RoboDK station: first project.rdk

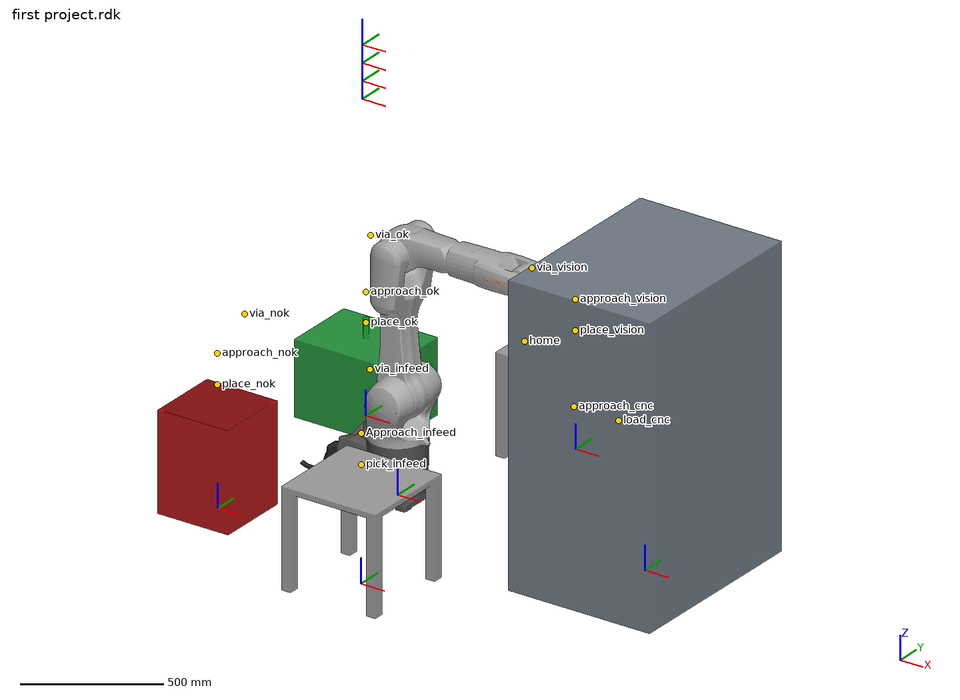
[picture v0: the station drawn from its stored meshes, robots at their saved joint values, targets as dots, program paths as lines]
Station KUKA_Cell (saved by RoboDK 6.1.1). Poses are relative to the parent item; angles as X-Y-Z fixed-axis rotations.
  - frame KUKA KR 10 R1100-2 Base at (0, 0, 0) mm
    - robot KUKA KR 10 R1100-2: 6 axes, payload 10.9 kg, reach 1101 mm, repeatability 0.02 mm, weight 56.5 kg
        modified DH rows (alpha deg, a mm, theta deg, d mm): 0, 0, 0, 400; -90, 25, 0, 0; 0, 560, -90, 0; -90, 25, 0, 515; 90, 0, 0, 0; -90, 0, 180, 90
        joint limits [-170, -190, -120, -185, -120, -350] to [170, 45, 156, 185, 120, 350]; home [0, -90, 90, 0, 0, 0]; saved at [0, -90, 90, 0, 90, 0]
      - tool Tool_Gripper, TCP at (0, 0, 150) mm, size 90 x 80 x 150 mm
    - target home (joint target) at (540, 0, 745) mm, rotated rx 180 ry 0 rz -180 deg; joints [0, -90, 90, 0, 90, 0] of KUKA KR 10 R1100-2
    - target via_infeed (joint target) at (226.29, -490.3, 745) mm, rotated rx 180 ry 0 rz 114.78 deg; joints [65.225, -90, 90, 0, 90, 0] of KUKA KR 10 R1100-2
    - target via_cnc (joint target) at (540, 0, 745) mm, rotated rx 180 ry 0 rz -180 deg; joints [0, -90, 90, 0, 90, 0] of KUKA KR 10 R1100-2
    - target via_vision (joint target) at (226.29, 490.3, 745) mm, rotated rx 180 ry 0 rz -114.78 deg; joints [-65.225, -90, 90, 0, 90, 0] of KUKA KR 10 R1100-2
    - target via_ok (joint target) at (-381.84, 381.84, 745) mm, rotated rx 180 ry 0 rz -45 deg; joints [-135, -90, 90, 0, 90, 0] of KUKA KR 10 R1100-2
    - target via_nok (joint target) at (-381.84, -381.84, 745) mm, rotated rx 180 ry 0 rz 45 deg; joints [135, -90, 90, 0, 90, 0] of KUKA KR 10 R1100-2
  - Python program check_paths (listed below)
  - Python program main_cycle (1) (listed below)
  - Python program build_cell (1) (listed below)
  - frame Frame_Infeed at (300, -650, 0) mm
    - object Table_Infeed at (0, 0, 0) mm, size 400 x 400 x 400 mm, geometry from Table.stl
    - target Approach_infeed (Cartesian target) at (0, 0, 580) mm, rotated rx 180 ry 0 rz 0 deg; joints [65.225, -70.524, 85.389, 0, 75.135, -114.775] of KUKA KR 10 R1100-2
    - target pick_infeed (Cartesian target) at (0, 0, 460) mm, rotated rx 180 ry 0 rz 0 deg; joints [65.225, -66.659, 93.982, 0, 62.678, -114.775] of KUKA KR 10 R1100-2
  - frame Frame_CNC at (1050, 0, 0) mm
    - object CNC_Machine at (0, 0, 0) mm, size 600 x 800 x 1200 mm, geometry from CNC_Machine.stl
    - target approach_cnc (Cartesian target) at (-300, 0, 550) mm, rotated rx 0 ry 90 rz 0 deg; joints [0, -74.689, 126.636, 0, -51.947, 0] of KUKA KR 10 R1100-2
    - target load_cnc (Cartesian target) at (-110, 0, 550) mm, rotated rx 0 ry 90 rz 0 deg; joints [0, -59.76, 102.885, 0, -43.124, 0] of KUKA KR 10 R1100-2
  - frame Frame_Vision at (300, 650, 0) mm
    - object Table_Vision at (0, 0, 0) mm, size 400 x 400 x 400 mm, geometry from Table.stl
    - target approach_vision (Cartesian target) at (0, 0, 580) mm, rotated rx 180 ry 0 rz 0 deg; joints [-65.225, -70.524, 85.389, 0, 75.135, 114.775] of KUKA KR 10 R1100-2
    - target place_vision (Cartesian target) at (0, 0, 460) mm, rotated rx 180 ry 0 rz 0 deg; joints [-65.225, -66.659, 93.982, 0, 62.678, 114.775] of KUKA KR 10 R1100-2
  - frame Frame_OK at (-450, 450, 0) mm
    - object Pallet_OK at (0, 0, 0) mm, size 400 x 300 x 300 mm, geometry from Pallet_OK.stl
    - target approach_ok (Cartesian target) at (0, 0, 480) mm, rotated rx 180 ry 0 rz 0 deg; joints [-135, -74.946, 103.078, 0, 61.868, 45] of KUKA KR 10 R1100-2
    - target place_ok (Cartesian target) at (0, 0, 360) mm, rotated rx 180 ry 0 rz 0 deg; joints [-135, -68.275, 109.448, 0, 48.827, 45] of KUKA KR 10 R1100-2
    - object Part_Shaft at (0, 0, 300) mm, size 20 x 20 x 80 mm, geometry from Part_Shaft.stl
  - frame Frame_NOK at (-450, -450, 0) mm
    - object Bin_NOK at (0, 0, 0) mm, size 300 x 300 x 400 mm, geometry from Bin_NOK.stl
    - target approach_nok (Cartesian target) at (0, 0, 600) mm, rotated rx 180 ry 0 rz 0 deg; joints [135, -78.926, 93.974, 0, 74.951, -45] of KUKA KR 10 R1100-2
    - target place_nok (Cartesian target) at (0, 0, 480) mm, rotated rx 180 ry 0 rz 0 deg; joints [135, -74.946, 103.078, 0, 61.868, -45] of KUKA KR 10 R1100-2
  - Python program kpi_report (listed below)
  - Python program dashboard (listed below)
  - frame HMI | ORDER OF-20261010-1825: 5 parts  |  now: SN-0005 at (-150, 0, 1700) mm
  - frame HMI | Status: ORDER FINISHED at (-150, 0, 1630) mm
  - frame HMI | Last: SN-0005  D=20.005 mm  OK  11.5 s  stop 152 s at (-150, 0, 1560) mm
  - frame HMI | Done 5/5   OK: 5   NOK: 0   Yield: 100 %   Downtime: 240 s at (-150, 0, 1490) mm

--- Python program check_paths ---
# =====================================================================
#  check_paths.py  -  checks every robot move of the cycle
#
#  For each move it checks:
#    1. REACH      : the robot can reach the target
#    2. COLLISION  : no collision along the path (robot / gripper vs cell)
#    3. LINEAR     : the straight-line (LIN) move is possible
#    4. SINGULARITY: wrist A5 not close to 0 deg (KUKA wrist singularity)
#    5. JOINT LIMIT: no joint closer than 5 deg to its limit
#
#  Run main_cycle.py at least once before (it writes the target values).
#  Result: a report in RoboDK + path_check_report.csv next to the station.
# =====================================================================
import csv
import os

from robodk.robolink import (Robolink, ITEM_TYPE_ROBOT, ITEM_TYPE_TOOL, ITEM_TYPE_TARGET,
                             ITEM_TYPE_FRAME, ITEM_TYPE_OBJECT, COLLISION_ON, COLLISION_OFF)
from robodk.robomath import transl

RDK = Robolink()

SIM_SPEED = 1          # 1 = real speed (slow, easy to watch). 5 = faster
SINGULARITY_DEG = 10   # warn if |A5| below this
LIMIT_MARGIN_DEG = 5   # warn if a joint is this close to its limit
HOME_JOINTS = [0, -90, 90, 0, 90, 0]

def find_robot_and_tool():
    """KUKA robot (ignores a gripper mechanism) + its gripper tool."""
    robots = RDK.ItemList(ITEM_TYPE_ROBOT)
    if not robots:
        raise Exception("No robot in the station. Load the KUKA KR 10 first.")
    rob = next((r for r in robots if "KUKA" in r.Name().upper()), robots[0])
    tl = RDK.Item('Tool_Gripper', ITEM_TYPE_TOOL)
    if not tl.Valid() or tl.Name() != 'Tool_Gripper':
        tools = [t for t in RDK.ItemList(ITEM_TYPE_TOOL)]
        if not tools:
            tl = rob.AddTool(transl(0, 0, 150), 'Tool_Gripper')
        else:
            tl = tools[0]
            tl.setName('Tool_Gripper')
    return rob, tl


robot, tool = find_robot_and_tool()
part = RDK.Item('Part_Shaft', ITEM_TYPE_OBJECT)
robot.setPoseTool(tool)


def collision_report():
    """Names of the items that are touching right now (empty string if none)."""
    try:
        pairs = RDK.CollisionPairs()            # [[item1, item2, link1, link2], ...]
        out = []
        for p in pairs:
            a = p[0].Name() + (f" (J{p[2]})" if len(p) > 2 and p[0].Type() == ITEM_TYPE_ROBOT else "")
            b = p[1].Name() + (f" (J{p[3]})" if len(p) > 3 and p[1].Type() == ITEM_TYPE_ROBOT else "")
            out.append(f"{a}  <->  {b}")
        return "; ".join(out)
    except Exception:
        try:
            return ", ".join(i.Name() for i in RDK.CollisionItems())
        except Exception:
            return ""


def choose_home():
    """Pick the home where the gripper points DOWN (A5 = +90 or -90).
    A home with the gripper pointing up makes the wrist flip during the moves
    and the gripper fingers hit the robot arm (self-collision)."""
    global HOME_JOINTS
    for a5 in (90, -90):
        j = [0, -90, 90, 0, a5, 0]
        robot.setJoints(j)
        tcp = robot.Pose()                  # TCP pose (active tool) in robot base
        if tcp[2, 2] < -0.5:                # tool Z axis points down
            HOME_JOINTS = j
            print(f"Home: A5 = {a5} (gripper pointing down)")
            return j
    return HOME_JOINTS

# Same sequence as main_cycle (OK branch + NOK branch)
SEQUENCE = [
    ("J", "home"),
    ("J", "via_infeed"), ("J", "Approach_infeed"), ("L", "pick_infeed"), ("GRIP", None),
    ("L", "Approach_infeed"), ("J", "via_infeed"),
    ("J", "via_cnc"), ("J", "approach_cnc"), ("L", "load_cnc"), ("RELEASE", "Frame_CNC"),
    ("L", "approach_cnc"), ("L", "load_cnc"), ("GRIP", None), ("L", "approach_cnc"), ("J", "via_cnc"),
    ("J", "via_vision"), ("J", "approach_vision"), ("L", "place_vision"), ("RELEASE", "Frame_Vision"),
    ("L", "approach_vision"), ("L", "place_vision"), ("GRIP", None), ("L", "approach_vision"),
    ("J", "via_vision"),
    ("J", "via_ok"), ("J", "approach_ok"), ("L", "place_ok"), ("RELEASE", "Frame_OK"),
    ("L", "approach_ok"), ("J", "via_ok"),
    ("J", "via_nok"), ("J", "approach_nok"), ("L", "place_nok"), ("L", "approach_nok"),  # NOK (empty gripper)
    ("J", "via_nok"),
    ("J", "home"),
]


def item(name, itype):
    it = RDK.Item(name, itype)
    if not it.Valid():
        raise Exception(f"Not found in the tree: {name}")
    return it


def disable_part_collisions():
    """The part touches the gripper and tables on purpose -> ignore it."""
    for other in RDK.ItemList():
        for link in range(8):
            try:
                RDK.setCollisionActivePair(COLLISION_OFF, part, other, 0, link)
            except Exception:
                pass


def as_list(values):
    """RoboDK returns joints as a Mat object -> convert to a flat Python list."""
    if hasattr(values, "rows"):          # robodk Mat (column or row vector)
        values = values.rows
    elif hasattr(values, "list"):
        values = values.list()
    out = []
    for v in values:
        if isinstance(v, (list, tuple)):
            out.extend(v)
        else:
            out.append(v)
    return [float(x) for x in out]


def check_joints(joints):
    """Return a list of warnings for singularity and joint limits."""
    warnings = []
    j = as_list(joints)
    if len(j) < 6:
        return warnings
    if abs(j[4]) < SINGULARITY_DEG:
        warnings.append(f"A5={j[4]:.1f} deg (near singularity)")
    limits = robot.JointLimits()
    lower, upper = as_list(limits[0]), as_list(limits[1])
    for i in range(6):
        if j[i] - lower[i] < LIMIT_MARGIN_DEG or upper[i] - j[i] < LIMIT_MARGIN_DEG:
            warnings.append(f"A{i+1}={j[i]:.1f} deg (near limit)")
    return warnings


# ---------------------------------------------------------------- run
RDK.setSimulationSpeed(SIM_SPEED)
RDK.setCollisionActive(COLLISION_ON)
disable_part_collisions()

part.setParent(item('Frame_Infeed', ITEM_TYPE_FRAME))
part.setPose(transl(0, 0, 400))
via = RDK.Item('via_infeed', ITEM_TYPE_TARGET)
if not via.Valid() or via.Name() != 'via_infeed':
    raise Exception('Run main_cycle once first (it creates the via_ points).')
robot.setJoints(item('home', ITEM_TYPE_TARGET).Joints())

report = []
n_problems = 0

for step, (kind, name) in enumerate(SEQUENCE, start=1):
    if kind == "GRIP":
        part.setParentStatic(tool)
        continue
    if kind == "RELEASE":
        part.setParentStatic(item(name, ITEM_TYPE_FRAME))
        continue

    target = item(name, ITEM_TYPE_TARGET)
    j_start = robot.Joints()
    row = {"step": step, "move": "PTP" if kind == "J" else "LIN", "target": name,
           "reach": "OK", "linear": "-", "collisions": 0, "hit": "", "warnings": "", "status": "OK"}

    # Test LIN feasibility before moving
    if kind == "L":
        robot.setPoseFrame(target.Parent())
        res = robot.MoveL_Test(j_start, target.Pose())
        row["linear"] = "OK" if res == 0 else ("collision" if res > 0 else "NOT POSSIBLE")

    # Execute the move (PTP if LIN impossible, like main_cycle does)
    try:
        if kind == "L" and row["linear"] != "NOT POSSIBLE":
            robot.MoveL(target)
        else:
            robot.MoveJ(target.Joints())     # joints computed by main_cycle setup
    except Exception:
        row["reach"] = "STOPPED (collision or unreachable)"
        row["hit"] = collision_report()
        row["status"] = "FAIL"
        report.append(row)
        n_problems += 1
        print(f"{step:02d} {name:16s} STOPPED (collision or unreachable)")
        break

    j_end = robot.Joints()
    # Collision along the joint path (PTP) or at the end pose
    if kind == "J":
        row["collisions"] = max(0, robot.MoveJ_Test(j_start, j_end))
    else:
        row["collisions"] = max(0, RDK.Collisions())
    if row["collisions"] > 0:
        row["hit"] = collision_report()
    warnings = check_joints(j_end)
    row["warnings"] = "; ".join(warnings)

    if row["collisions"] > 0 or row["linear"] in ("collision", "NOT POSSIBLE"):
        row["status"] = "FAIL"
    elif warnings:
        row["status"] = "WARNING"
    if row["status"] != "OK":
        n_problems += 1

    report.append(row)
    print(f"{step:02d} {row['move']} {name:16s} reach={row['reach']:4s} "
          f"lin={row['linear']:12s} coll={row['collisions']} {row['status']} {row['warnings']}")

RDK.setCollisionActive(COLLISION_OFF)

# ---------------------------------------------------------------- report
station_path = RDK.getParam('PATH_OPENSTATION')
out_dir = station_path if station_path and os.path.isdir(station_path) else os.path.expanduser("~")
out_file = os.path.join(out_dir, "path_check_report.csv")
with open(out_file, "w", newline="") as f:
    w = csv.DictWriter(f, fieldnames=list(report[0].keys()))
    w.writeheader()
    w.writerows(report)

lines = [f"{r['step']:02d} {r['move']} {r['target']}: {r['status']}"
         + (f" {r['reach']}" if r['reach'] != 'OK' else "")
         + (f" ({r['warnings']})" if r['warnings'] else "")
         + (f" collisions={r['collisions']}" if r['collisions'] else "")
         + (f"\n      HIT: {r['hit']}" if r['hit'] else "")
         + (f" LIN={r['linear']}" if r['linear'] not in ('-', 'OK') else "")
         for r in report]
summary = ("ALL PATHS OK" if n_problems == 0 else f"{n_problems} PROBLEM(S) FOUND")
RDK.ShowMessage(summary + "\n\n" + "\n".join(lines) + f"\n\nReport: {out_file}", True)
print(summary, "->", out_file)

--- Python program main_cycle (1) ---
# =====================================================================
#  KUKA KR 10 machine-tending cell - main cycle (RoboDK Python API)
#
#  1. SETUP : writes every target, picks ONE consistent arm configuration
#             per station (no wrist flips) and creates a safe "via" point
#             above each station.
#  2. CYCLE : pick -> CNC -> vision -> OK / NOK, always moving between
#             stations at safe height (via points).
#  3. LOG   : one CSV line per part (for the MES dashboard).
#
#  Tip: run it once with collision checking OFF (setup), then check_paths.
# =====================================================================
import csv
import math
import os
import random
import time
from datetime import datetime

from robodk.robolink import (Robolink, ITEM_TYPE_ROBOT, ITEM_TYPE_TOOL,
                             ITEM_TYPE_TARGET, ITEM_TYPE_FRAME, ITEM_TYPE_OBJECT,
                             COLLISION_ON, COLLISION_OFF)
from robodk.robomath import transl, invH, KUKA_2_Pose

RDK = Robolink()

# ---------------------------------------------------------------- settings
N_PARTS = 5                      # number of parts to produce
MACHINING_TIME_S = 3             # simulated CNC cycle
NOMINAL_DIAM = 20.00             # mm
TOLERANCE = 0.05                 # mm  -> OK if 19.95 .. 20.05
_station_dir = RDK.getParam('PATH_OPENSTATION')          # folder of the saved station
LOG_DIR = _station_dir if _station_dir and os.path.isdir(str(_station_dir)) else \
    os.path.join(os.path.expanduser("~"), "Documents", "KUKA_Cell_MES")
LOG_FILE = os.path.join(LOG_DIR, "kuka_cell_log.csv")   # CSV saved next to KUKA_Cell.rdk
CNC_FRAME_X = 1050               # CNC farther: more space between robot and CNC door

# ---------------------------------------------------------------- STEP 1: faults & downtime
# Each fault: (station, stop reason, probability per part, min-max stop duration in seconds)
FAULTS = [
    ("infeed", "Part missing on infeed",   0.10, (20, 60)),
    ("infeed", "Gripper fault",            0.05, (30, 90)),
    ("cnc",    "CNC door not open",        0.08, (15, 45)),
    ("cnc",    "Tool change on CNC",       0.05, (60, 180)),
    ("vision", "Camera timeout",           0.07, (10, 30)),
]
TIME_SCALE = 0.05                # a 60 s stop is shown as 3 s in the simulation
EVENT_FILE = os.path.join(LOG_DIR, "kuka_cell_events.csv")   # one line per stop
ORDER_ID = datetime.now().strftime("OF-%Y%m%d-%H%M")         # production order number

# Stations: name -> (frame, approach target, work target, approach values, work values)
# values = (X, Y, Z, A=rz, B=ry, C=rx) in the station frame (KUKA convention)
STATIONS = {
    "infeed": ("Frame_Infeed", "Approach_infeed", "pick_infeed",
               (0, 0, 580, 0, 0, 180), (0, 0, 460, 0, 0, 180)),
    "cnc":    ("Frame_CNC", "approach_cnc", "load_cnc",
               (-300, 0, 550, 0, 90, 0), (-110, 0, 550, 0, 90, 0)),
    "vision": ("Frame_Vision", "approach_vision", "place_vision",
               (0, 0, 580, 0, 0, 180), (0, 0, 460, 0, 0, 180)),
    "ok":     ("Frame_OK", "approach_ok", "place_ok",
               (0, 0, 480, 0, 0, 180), (0, 0, 360, 0, 0, 180)),
    "nok":    ("Frame_NOK", "approach_nok", "place_nok",
               (0, 0, 600, 0, 0, 180), (0, 0, 480, 0, 0, 180)),
}
HOME_JOINTS = [0, -90, 90, 0, 90, 0]
SOLVED = {}        # target name -> joints computed in setup (used by MoveJ)

# ---------------------------------------------------------------- items
def find_robot_and_tool():
    """KUKA robot (ignores a gripper mechanism) + its gripper tool."""
    robots = RDK.ItemList(ITEM_TYPE_ROBOT)
    if not robots:
        raise Exception("No robot in the station. Load the KUKA KR 10 first.")
    rob = next((r for r in robots if "KUKA" in r.Name().upper()), robots[0])
    tl = RDK.Item('Tool_Gripper', ITEM_TYPE_TOOL)
    if not tl.Valid() or tl.Name() != 'Tool_Gripper':
        tools = [t for t in RDK.ItemList(ITEM_TYPE_TOOL)]
        if not tools:
            tl = rob.AddTool(transl(0, 0, 150), 'Tool_Gripper')
        else:
            tl = tools[0]
            tl.setName('Tool_Gripper')
    return rob, tl


robot, tool = find_robot_and_tool()
part = RDK.Item('Part_Shaft', ITEM_TYPE_OBJECT)
robot.setPoseTool(tool)


def collision_report():
    """Names of the items that are touching right now (empty string if none)."""
    try:
        pairs = RDK.CollisionPairs()            # [[item1, item2, link1, link2], ...]
        out = []
        for p in pairs:
            a = p[0].Name() + (f" (J{p[2]})" if len(p) > 2 and p[0].Type() == ITEM_TYPE_ROBOT else "")
            b = p[1].Name() + (f" (J{p[3]})" if len(p) > 3 and p[1].Type() == ITEM_TYPE_ROBOT else "")
            out.append(f"{a}  <->  {b}")
        return "; ".join(out)
    except Exception:
        try:
            return ", ".join(i.Name() for i in RDK.CollisionItems())
        except Exception:
            return ""
robot.setPoseFrame(robot.Parent())      # poses measured in the robot base


def T(name):
    item = RDK.Item(name, ITEM_TYPE_TARGET)
    if not item.Valid() or item.Name() != name:
        raise Exception(f"Target not found in the tree: {name}")
    return item


def F(name):
    item = RDK.Item(name, ITEM_TYPE_FRAME)
    if not item.Valid():
        raise Exception(f"Frame not found in the tree: {name}")
    return item


def as_list(values):
    """RoboDK returns joints as a Mat -> flat Python list."""
    if hasattr(values, "rows"):
        values = values.rows
    elif hasattr(values, "list"):
        values = values.list()
    out = []
    for v in values:
        out.extend(v) if isinstance(v, (list, tuple)) else out.append(v)
    return [float(x) for x in out]


# ---------------------------------------------------------------- moves
def MJ(name):
    try:
        if name in SOLVED:
            robot.MoveJ(SOLVED[name])        # exact joints from setup: no config surprise
        else:
            robot.MoveJ(T(name))
    except Exception as e:
        hit = collision_report()
        msg = f"Move stopped going to: {name}" + (f"\nCOLLISION: {hit}" if hit else f" ({e})")
        RDK.ShowMessage(msg, True)
        raise Exception(msg)


def ML(name):
    try:
        robot.MoveL(T(name))
    except Exception:
        print(f"  MoveL to {name} not possible -> MoveJ used")
        MJ(name)


def grip():
    part.setParentStatic(tool)


def release(frame_name):
    part.setParentStatic(F(frame_name))


# ---------------------------------------------------------------- on-screen display (HMI)
# RoboDK shows the NAME of a frame as a text label in the 3D view.
# We create 4 small frames above the cell and change their names = live text panel.
HMI_POS = (-150, 0, 1700)          # where the text panel floats (mm, station frame)
HMI = []
PART_COLOR = [0.85, 0.65, 0.20, 1]   # gold = raw part


def hmi_init():
    for fr in RDK.ItemList(ITEM_TYPE_FRAME):          # remove the panel of a previous run
        if fr.Name().startswith("HMI"):
            fr.Delete()
    HMI.clear()
    for i in range(4):
        fr = RDK.AddFrame(f"HMI {i}")
        fr.setPose(transl(HMI_POS[0], HMI_POS[1], HMI_POS[2] - 70 * i))
        try:
            fr.setVisible(True, False)                  # show the text, hide the axes
        except Exception:
            pass
        HMI.append(fr)


def hmi(line, text):
    """Write one line of the 3D text panel (0 = title, 1 = status, 2 = last part, 3 = totals)."""
    if line < len(HMI):
        HMI[line].setName(f"HMI | {text}")


def color_part(rgba):
    try:
        part.setColor(rgba)
    except Exception:
        pass


def reset_part():
    part.setParent(F('Frame_Infeed'))
    part.setPose(transl(0, 0, 400))
    color_part(PART_COLOR)


# ---------------------------------------------------------------- setup helpers
def choose_home():
    """Home with the gripper pointing DOWN (A5 = +90 or -90)."""
    global HOME_JOINTS
    for a5 in (90, -90):
        j = [0, -90, 90, 0, a5, 0]
        robot.setJoints(j)
        if robot.Pose()[2, 2] < -0.5:        # tool Z axis points down
            HOME_JOINTS = j
            break
    print(f"Home joints: {HOME_JOINTS}")


def get_or_create_target(name, parent):
    item = RDK.Item(name, ITEM_TYPE_TARGET)
    if not item.Valid() or item.Name() != name:
        item = RDK.AddTarget(name, parent, robot)
    item.setParent(parent)
    return item


def via_joints(frame_name):
    """Home posture rotated (A1) toward the station: high and safe."""
    p = F(frame_name).PoseAbs().Pos()
    best, best_dot = None, -2
    ang = math.degrees(math.atan2(p[1], p[0]))
    for a1 in (ang, -ang):
        j = list(HOME_JOINTS)
        j[0] = a1
        robot.setJoints(j)
        t = robot.Pose().Pos()
        n = math.hypot(t[0], t[1]) * math.hypot(p[0], p[1]) or 1
        dot = (t[0] * p[0] + t[1] * p[1]) / n
        if dot > best_dot:
            best, best_dot = j, dot
    return best


def flange_pose(frame_name, values):
    """Flange pose in the robot base for a TCP target given in a station frame."""
    base_abs = robot.Parent().PoseAbs()
    frame_abs = F(frame_name).PoseAbs()
    return invH(base_abs) * frame_abs * KUKA_2_Pose(list(values)) * invH(robot.PoseTool())


def ik(frame_name, values, joints_approx):
    target = flange_pose(frame_name, values)
    sol = as_list(robot.SolveIK(target, joints_approx))
    if len(sol) < 6:
        return None
    sol = sol[:6]
    # verify: forward kinematics must give back the same flange position
    fk = robot.SolveFK(sol)
    err = sum((a - b) ** 2 for a, b in zip(fk.Pos(), target.Pos())) ** 0.5
    if err > 1.0:
        return None
    lower, upper = [as_list(x) for x in robot.JointLimits()[:2]]
    if any(not (lo <= v <= up) for v, lo, up in zip(sol, lower, upper)):
        return None
    return sol


def path_free(j_from, j_to, frame_name=None, work_values=None):
    """True if the PTP move j_from->j_to (and the LIN to the work point) is collision free."""
    try:
        if robot.MoveJ_Test(j_from, j_to) != 0:
            return False
        robot.setJoints(j_to)
        if RDK.Collisions() > 0:
            return False
        if frame_name and work_values:
            robot.setPoseFrame(F(frame_name))
            res = robot.MoveL_Test(j_to, KUKA_2_Pose(list(work_values)))
            robot.setPoseFrame(robot.Parent())
            if res != 0:
                return False
        return True
    except Exception:
        robot.setPoseFrame(robot.Parent())
        return True        # if the test itself is not available, do not block


def setup_cell():
    print("SETUP...")
    RDK.Render(False)
    RDK.setCollisionActive(COLLISION_ON)       # setup picks collision-free configurations
    F('Frame_CNC').setPose(transl(CNC_FRAME_X, 0, 0))
    choose_home()

    base = robot.Parent()
    home = get_or_create_target('home', base)
    home.setAsJointTarget()
    home.setJoints(HOME_JOINTS)
    SOLVED['home'] = list(HOME_JOINTS)

    for key, (frame, appr, work, v_appr, v_work) in STATIONS.items():
        # safe point above the station
        vj = via_joints(frame)
        via = get_or_create_target(f'via_{key}', base)
        via.setAsJointTarget()
        via.setJoints(vj)
        SOLVED[f'via_{key}'] = vj

        # approach + work: same wrist orientation, configuration close to the via point
        done = False
        candidates = [(extra, t, dz) for dz in (0, 100) for t in (0, 0.25, 0.5)
                      for extra in (0, 180, 90, -90)]
        for extra, t, dz in candidates:
            # approach can be moved a bit toward the work point if too far / too folded
            va = [a + t * (w - a) for a, w in zip(v_appr[:3], v_work[:3])] + list(v_appr[3:])
            va[5] += extra
            if key != "cnc":
                va[2] += dz                    # higher approach if needed (not for the CNC door)
            vw = list(v_work); vw[5] += extra
            ja = ik(frame, va, vj)
            jw = ik(frame, vw, ja) if ja else None
            if (ja and jw and abs(ja[0] - vj[0]) < 60 and abs(jw[4] - ja[4]) < 60
                    and path_free(vj, ja, frame, vw)):
                for name, vals, joints in ((appr, va, ja), (work, vw, jw)):
                    tgt = get_or_create_target(name, F(frame))
                    tgt.setAsCartesianTarget()
                    tgt.setPose(KUKA_2_Pose(vals))
                    tgt.setJoints(joints)    # stored configuration -> no wrist flip
                    SOLVED[name] = joints
                print(f"  {key:6s}: OK collision-free (wrist +{extra} deg, approach shifted {int(t*100)}%, +{dz} mm)")
                done = True
                break
        if not done:
            RDK.Render(True)
            p = F(frame).PoseAbs().Pos()
            raise Exception(f"Station {key}: no reachable AND collision-free configuration. "
                            f"Frame at X={p[0]:.0f} Y={p[1]:.0f}. Tell Claude this message.")

    # check the moves between stations (home -> via -> via ...)
    order = ['home', 'via_infeed', 'via_cnc', 'via_vision', 'via_ok', 'via_vision', 'via_nok', 'home']
    for a, b in zip(order, order[1:]):
        if robot.MoveJ_Test(SOLVED[a], SOLVED[b]) != 0:
            print(f"  WARNING: collision on the move {a} -> {b}: {collision_report()}")

    robot.setJoints(HOME_JOINTS)
    RDK.Render(True)
    print("SETUP done.\n")


# ---------------------------------------------------------------- cycle
def go_station(key):
    MJ(f'via_{key}')
    MJ(STATIONS[key][1])           # approach


def leave_station(key):
    ML(STATIONS[key][1])           # back to approach
    MJ(f'via_{key}')


def write_csv(path, row):
    """Append one row to a CSV file (header written the first time).
    If an old file has different columns, it is renamed *_old.csv."""
    os.makedirs(os.path.dirname(path), exist_ok=True)
    if os.path.exists(path):
        with open(path, newline="") as f:
            header = f.readline().strip().split(",")
        if header != list(row.keys()):
            os.replace(path, path.replace(".csv", "_old.csv"))
    new_file = not os.path.exists(path)
    with open(path, "a", newline="") as f:
        w = csv.DictWriter(f, fieldnames=list(row.keys()))
        if new_file:
            w.writeheader()
        w.writerow(row)


def check_faults(serial, station):
    """Random stops at a station. Returns the downtime (s) and the wait time used."""
    downtime, waited = 0.0, 0.0
    for st, reason, prob, (dmin, dmax) in FAULTS:
        if st == station and random.random() < prob:
            duration = random.uniform(dmin, dmax)
            start = datetime.now()
            hmi(1, f"Status: FAULT - {reason} ({duration:.0f} s)")
            RDK.ShowMessage(f"FAULT at {station}: {reason}", False)
            wait = duration * TIME_SCALE
            time.sleep(wait)
            write_csv(EVENT_FILE, {
                "order": ORDER_ID,
                "serial": serial,
                "station": station,
                "reason": reason,
                "start": start.isoformat(timespec="seconds"),
                "duration_s": round(duration, 1),
            })
            downtime += duration
            waited += wait
    return downtime, waited


def run_cycle(serial):
    t0 = time.time()
    downtime, waited = 0.0, 0.0
    hmi(0, f"ORDER {ORDER_ID}: {N_PARTS} parts  |  now: {serial}")
    reset_part()
    MJ('home')

    # PICK
    hmi(1, "Status: PICKING raw part")
    d, w = check_faults(serial, "infeed"); downtime += d; waited += w
    hmi(1, "Status: PICKING raw part")
    go_station('infeed')
    ML('pick_infeed')
    grip()
    leave_station('infeed')

    # CNC load / machining / unload
    hmi(1, "Status: LOADING CNC")
    d, w = check_faults(serial, "cnc"); downtime += d; waited += w
    hmi(1, "Status: LOADING CNC")
    go_station('cnc')
    ML('load_cnc')
    release('Frame_CNC')
    ML('approach_cnc')
    hmi(1, f"Status: MACHINING ({MACHINING_TIME_S} s)")
    time.sleep(MACHINING_TIME_S)
    hmi(1, "Status: UNLOADING CNC")
    ML('load_cnc')
    grip()
    leave_station('cnc')

    # VISION
    hmi(1, "Status: VISION INSPECTION")
    d, w = check_faults(serial, "vision"); downtime += d; waited += w
    hmi(1, "Status: VISION INSPECTION")
    go_station('vision')
    ML('place_vision')
    release('Frame_Vision')
    ML('approach_vision')
    diameter = random.gauss(NOMINAL_DIAM, 0.02)
    ok = abs(diameter - NOMINAL_DIAM) <= TOLERANCE
    color_part([0.1, 0.8, 0.2, 1] if ok else [0.9, 0.1, 0.1, 1])     # green OK / red NOK
    hmi(1, f"Status: MEASURED D={diameter:.3f} mm -> {'OK' if ok else 'NOK'}")
    time.sleep(1)
    ML('place_vision')
    grip()
    leave_station('vision')

    # OK pallet or NOK bin
    hmi(1, f"Status: SORTING to {'OK pallet' if ok else 'NOK bin'}")
    key = 'ok' if ok else 'nok'
    go_station(key)
    ML(STATIONS[key][2])
    release(STATIONS[key][0])
    leave_station(key)
    MJ('home')

    return {"order": ORDER_ID,
            "timestamp": datetime.now().isoformat(timespec="seconds"),
            "serial": serial,
            "diameter_mm": round(diameter, 3),
            "result": 'OK' if ok else 'NOK',
            "cycle_time_s": round(time.time() - t0 - waited, 1),   # running time only
            "downtime_s": round(downtime, 1)}                       # stops (real seconds)


def log_row(row):
    write_csv(LOG_FILE, row)


# ---------------------------------------------------------------- main
setup_cell()
hmi_init()
hmi(0, f"ORDER: {N_PARTS} parts  |  tolerance {NOMINAL_DIAM:.2f} +/- {TOLERANCE} mm")
hmi(1, "Status: READY")
hmi(2, "Last part: -")
hmi(3, "OK: 0   NOK: 0")

n_ok = 0
for i in range(1, N_PARTS + 1):
    row = run_cycle(f"SN-{i:04d}")
    log_row(row)
    n_ok += row["result"] == "OK"
    msg = (f"{row['serial']} | diam={row['diameter_mm']} mm | "
           f"{row['result']} | cycle={row['cycle_time_s']} s")
    print(msg)
    RDK.ShowMessage(msg, False)
    done = i
    total_down = globals().get("total_down", 0) + row["downtime_s"]
    globals()["total_down"] = total_down
    hmi(2, f"Last: {row['serial']}  D={row['diameter_mm']} mm  {row['result']}  "
           f"{row['cycle_time_s']} s  stop {row['downtime_s']:.0f} s")
    hmi(3, f"Done {done}/{N_PARTS}   OK: {n_ok}   NOK: {done - n_ok}   "
           f"Yield: {100 * n_ok / done:.0f} %   Downtime: {total_down:.0f} s")

summary = f"DONE: {N_PARTS} parts, {n_ok} OK, {N_PARTS - n_ok} NOK. Log: {LOG_FILE}"
print(summary)
RDK.ShowMessage(summary, False)
hmi(1, "Status: ORDER FINISHED")

--- Python program build_cell (1) ---
# =====================================================================
#  build_cell.py  -  builds the whole KUKA cell automatically in RoboDK
#
#  Before running:
#   - The station must already contain: KUKA KR 10 R1100-2 + RobotiQ gripper
#     + a tool named "Tool_Gripper" (TCP Z = 150).
#   - Unzip KUKA_Cell_Models.zip anywhere (Downloads, Documents, Desktop...)
#
#  Run it once (Python program in RoboDK -> double-click).
#  It creates frames, objects, targets, then SAVES the station
#  as KUKA_Cell.rdk next to the STL files.
#  Then run main_cycle.py to produce parts.
# =====================================================================
import os

from robodk.robolink import (Robolink, ITEM_TYPE_ROBOT, ITEM_TYPE_TOOL,
                             ITEM_TYPE_FRAME, ITEM_TYPE_OBJECT, ITEM_TYPE_TARGET)
from robodk.robomath import transl, eye

RDK = Robolink()

NEEDED = ["Table.stl", "Part_Shaft.stl", "CNC_Machine.stl", "Pallet_OK.stl", "Bin_NOK.stl"]


def find_models_dir():
    """Look for the folder that contains the 5 STL files (Documents, OneDrive,
    Downloads, Desktop...). If not found, ask the user to pick the folder."""
    home = os.path.expanduser("~")
    roots = [os.path.join(home, d) for d in
             ("Documents", "OneDrive", "Downloads",
              "Desktop", "Bureau")]
    roots += [os.path.join(home, "OneDrive", d) for d in ("Documents", "Desktop", "Bureau")]
    roots += ["C:\\KUKA_Cell_MES"]
    for root in roots:
        if not os.path.isdir(root):
            continue
        base_depth = root.rstrip("\\/").count(os.sep)
        for folder, subdirs, files in os.walk(root):
            if folder.count(os.sep) - base_depth > 4:
                subdirs[:] = []          # don't search too deep
                continue
            if all(f in files for f in NEEDED):
                return folder
    # Not found automatically -> folder picker
    try:
        import tkinter
        from tkinter import filedialog
        win = tkinter.Tk()
        win.withdraw()
        win.attributes("-topmost", True)
        folder = filedialog.askdirectory(title="Select the folder that contains the 5 STL files")
        win.destroy()
        if folder and all(os.path.exists(os.path.join(folder, f)) for f in NEEDED):
            return folder
    except Exception:
        pass
    return None


MODELS_DIR = find_models_dir()
if MODELS_DIR is None:
    raise Exception("The 5 STL files were not found. Unzip KUKA_Cell_Models.zip "
                    "into Documents\\KUKA_Cell_MES\\models and run again.")
# Project folder = the folder above "models" (or the models folder itself)
PROJECT_DIR = (os.path.dirname(MODELS_DIR)
               if os.path.basename(MODELS_DIR).lower() == "models" else MODELS_DIR)
STATION_FILE = os.path.join(PROJECT_DIR, "KUKA_Cell.rdk")
print(f"Models found in: {MODELS_DIR}")

# Frames: name -> (X, Y, Z) relative to the station
FRAMES = {
    "Frame_Infeed": (300, -650, 0),
    "Frame_CNC":    (1050, 0, 0),
    "Frame_Vision": (300, 650, 0),
    "Frame_OK":     (-450, 450, 0),
    "Frame_NOK":    (-450, -450, 0),
}

# Objects: name -> (STL file, frame, Z offset, color RGBA 0-1)
OBJECTS = {
    "Table_Infeed": ("Table.stl",       "Frame_Infeed", 0,   [0.75, 0.75, 0.75, 1]),
    "Part_Shaft":   ("Part_Shaft.stl",  "Frame_Infeed", 400, [0.85, 0.65, 0.20, 1]),
    "CNC_Machine":  ("CNC_Machine.stl", "Frame_CNC",    0,   [0.55, 0.60, 0.65, 1]),
    "Table_Vision": ("Table.stl",       "Frame_Vision", 0,   [0.75, 0.75, 0.75, 1]),
    "Pallet_OK":    ("Pallet_OK.stl",   "Frame_OK",     0,   [0.20, 0.70, 0.30, 1]),
    "Bin_NOK":      ("Bin_NOK.stl",     "Frame_NOK",    0,   [0.85, 0.15, 0.15, 1]),
}

# Targets: name -> frame (values are written later by main_cycle.py)
TARGETS = {
    "Approach_infeed": "Frame_Infeed", "pick_infeed": "Frame_Infeed",
    "approach_cnc": "Frame_CNC",       "load_cnc": "Frame_CNC",
    "approach_vision": "Frame_Vision", "place_vision": "Frame_Vision",
    "approach_ok": "Frame_OK",         "place_ok": "Frame_OK",
    "approach_nok": "Frame_NOK",       "place_nok": "Frame_NOK",
}
HOME_JOINTS = [0, -90, 90, 0, 90, 0]


def delete_if_exists(name, item_type):
    item = RDK.Item(name, item_type)
    while item.Valid() and item.Name() == name:
        item.Delete()
        item = RDK.Item(name, item_type)


# ---------------------------------------------------------------- checks
def find_robot_and_tool():
    """KUKA robot (ignores a gripper mechanism) + its gripper tool."""
    robots = RDK.ItemList(ITEM_TYPE_ROBOT)
    if not robots:
        raise Exception("No robot in the station. Load the KUKA KR 10 first.")
    rob = next((r for r in robots if "KUKA" in r.Name().upper()), robots[0])
    tl = RDK.Item('Tool_Gripper', ITEM_TYPE_TOOL)
    if not tl.Valid() or tl.Name() != 'Tool_Gripper':
        tools = [t for t in RDK.ItemList(ITEM_TYPE_TOOL)]
        if not tools:
            tl = rob.AddTool(transl(0, 0, 150), 'Tool_Gripper')
        else:
            tl = tools[0]
            tl.setName('Tool_Gripper')
    return rob, tl


robot, tool = find_robot_and_tool()

# ---------------------------------------------------------------- gripper
# Free license = max 1 robot: remove any gripper "mechanism" (counted as a robot)
for r in RDK.ItemList(ITEM_TYPE_ROBOT):
    if r.Name() != robot.Name():
        r.Delete()
for fr in RDK.ItemList(ITEM_TYPE_FRAME):
    if "ROBOTIQ" in fr.Name().upper():
        fr.Delete()
# Re-create the gripper tool with its 3D shape (Gripper_2F.stl)
for t in RDK.ItemList(ITEM_TYPE_TOOL):
    t.Delete()
tool = robot.AddTool(transl(0, 0, 150), 'Tool_Gripper')     # TCP between the fingertips
gripper_stl = os.path.join(MODELS_DIR, "Gripper_2F.stl")
if os.path.exists(gripper_stl):
    shape = RDK.AddFile(gripper_stl)
    tool.AddGeometry(shape, eye(4))
    shape.Delete()
    try:
        tool.setColor([0.15, 0.15, 0.15, 1])
    except Exception:
        pass
    print("Gripper  Gripper_2F.stl added on the robot flange")
else:
    print("WARNING: Gripper_2F.stl not found next to the other STL files -> tool without shape")
if not os.path.isdir(MODELS_DIR):
    raise Exception(f"Models folder not found: {MODELS_DIR}\n"
                    f"Unzip KUKA_Cell_Models.zip there.")

RDK.Render(False)

# Robot base at the origin of the station
robot.Parent().setPose(eye(4))
robot.setPoseTool(tool)

# ---------------------------------------------------------------- frames
frames = {}
for name, (x, y, z) in FRAMES.items():
    delete_if_exists(name, ITEM_TYPE_FRAME)   # also deletes its children
    fr = RDK.AddFrame(name)
    fr.setPose(transl(x, y, z))
    frames[name] = fr
    print(f"Frame   {name:14s} at ({x}, {y}, {z})")

# ---------------------------------------------------------------- objects
for name, (stl, frame, z, color) in OBJECTS.items():
    path = os.path.join(MODELS_DIR, stl)
    if not os.path.exists(path):
        raise Exception(f"Missing model file: {path}")
    obj = RDK.AddFile(path, frames[frame])
    obj.setName(name)
    obj.setPose(transl(0, 0, z))
    obj.setColor(color)
    print(f"Object  {name:14s} in {frame}")

# ---------------------------------------------------------------- targets
robot.setJoints(HOME_JOINTS)
delete_if_exists("home", ITEM_TYPE_TARGET)
home = RDK.AddTarget("home", robot.Parent(), robot)
home.setAsJointTarget()
home.setJoints(HOME_JOINTS)
print("Target  home (joints)")

for name, frame in TARGETS.items():
    tgt = RDK.AddTarget(name, frames[frame], robot)
    print(f"Target  {name:14s} in {frame}")

RDK.Render(True)

# ---------------------------------------------------------------- save
os.makedirs(PROJECT_DIR, exist_ok=True)
RDK.ActiveStation().setName("KUKA_Cell")
RDK.Save(STATION_FILE)
msg = f"Cell built and saved to {STATION_FILE}. Now run main_cycle.py"
print(msg)
RDK.ShowMessage(msg, False)

--- Python program kpi_report ---
# =====================================================================
#  kpi_report.py  -  STEP 2: computes the cell KPIs from the MES logs
#
#  Reads:   kuka_cell_log.csv     (one line per part)
#           kuka_cell_events.csv  (one line per stop)
#  Computes: OEE = Availability x Performance x Quality
#            yield, cycle times, MTBF, MTTR, downtime Pareto
#  Writes:  kpi_report.txt  (+ shows it in RoboDK if run from RoboDK)
#
#  Run it from RoboDK (Python program, double-click) or with: python kpi_report.py
# =====================================================================
import csv
import os
from collections import defaultdict

# ---------------------------------------------------------------- settings
ONLY_LAST_ORDER = True     # True = KPIs of the last production order only
IDEAL_CYCLE_S = None       # ideal cycle time (s). None = best cycle observed


# ---------------------------------------------------------------- find the files
def find_log_dir():
    candidates = []
    try:                                           # folder of the RoboDK station
        from robodk.robolink import Robolink
        d = Robolink().getParam('PATH_OPENSTATION')
        if d:
            candidates.append(str(d))
    except Exception:
        pass
    here = os.path.dirname(os.path.abspath(__file__))
    home = os.path.expanduser("~")
    candidates += [here, os.path.join(home, "Documents", "KUKA_Cell_MES")]
    for c in candidates:
        if os.path.exists(os.path.join(c, "kuka_cell_log.csv")):
            return c
    for root in [os.path.join(home, d) for d in ("Documents", "OneDrive", "Downloads", "Desktop")]:
        if not os.path.isdir(root):
            continue
        base = root.count(os.sep)
        for folder, subdirs, files in os.walk(root):
            if folder.count(os.sep) - base > 4:
                subdirs[:] = []
                continue
            if "kuka_cell_log.csv" in files:
                return folder
    raise Exception("kuka_cell_log.csv not found. Run main_cycle first.")


def read_csv(path):
    if not os.path.exists(path):
        return []
    with open(path, newline="") as f:
        return list(csv.DictReader(f))


# ---------------------------------------------------------------- KPI calculation
def compute(parts, events):
    n = len(parts)
    if n == 0:
        raise Exception("No parts in the log.")
    n_ok = sum(1 for p in parts if p["result"] == "OK")
    cycles = [float(p["cycle_time_s"]) for p in parts]
    run_time = sum(cycles)                                        # robot working
    downtime = sum(float(e["duration_s"]) for e in events)       # cell stopped
    planned = run_time + downtime                                # total production time
    ideal = IDEAL_CYCLE_S or min(cycles)

    availability = run_time / planned if planned else 0
    performance = min(1.0, ideal * n / run_time) if run_time else 0
    quality = n_ok / n
    oee = availability * performance * quality

    n_stops = len(events)
    mtbf = run_time / n_stops if n_stops else None              # mean time between failures
    mttr = downtime / n_stops if n_stops else None              # mean time to repair

    pareto = defaultdict(lambda: [0, 0.0])                      # reason -> [count, seconds]
    for e in events:
        pareto[e["reason"]][0] += 1
        pareto[e["reason"]][1] += float(e["duration_s"])
    pareto = sorted(pareto.items(), key=lambda kv: kv[1][1], reverse=True)

    return {
        "parts": n, "ok": n_ok, "nok": n - n_ok,
        "run_time": run_time, "downtime": downtime, "planned": planned,
        "ideal": ideal, "avg_cycle": run_time / n, "min_cycle": min(cycles), "max_cycle": max(cycles),
        "availability": availability, "performance": performance, "quality": quality, "oee": oee,
        "stops": n_stops, "mtbf": mtbf, "mttr": mttr, "pareto": pareto,
    }


def fmt_report(order, k):
    pct = lambda x: f"{100 * x:5.1f} %"
    sec = lambda x: "-" if x is None else f"{x:6.1f} s"
    lines = [
        f"KPI REPORT  -  order {order}",
        "=" * 46,
        f"Parts produced      : {k['parts']}   (OK {k['ok']} / NOK {k['nok']})",
        f"Planned time        : {k['planned']:.1f} s",
        f"Running time        : {k['run_time']:.1f} s",
        f"Downtime            : {k['downtime']:.1f} s  in {k['stops']} stops",
        "-" * 46,
        f"Availability (A)    : {pct(k['availability'])}   running / planned",
        f"Performance  (P)    : {pct(k['performance'])}   ideal x parts / running",
        f"Quality      (Q)    : {pct(k['quality'])}   OK / produced",
        f"OEE = A x P x Q     : {pct(k['oee'])}",
        "-" * 46,
        f"Cycle time avg/min/max : {k['avg_cycle']:.1f} / {k['min_cycle']:.1f} / {k['max_cycle']:.1f} s",
        f"Ideal cycle time       : {k['ideal']:.1f} s",
        f"MTBF (between stops)   : {sec(k['mtbf'])}",
        f"MTTR (repair time)     : {sec(k['mttr'])}",
        "-" * 46,
        "Downtime Pareto (biggest loss first):",
    ]
    for reason, (count, seconds) in k["pareto"]:
        share = seconds / k["downtime"] if k["downtime"] else 0
        lines.append(f"  {reason:26s} {count:2d}x  {seconds:6.1f} s  {pct(share)}")
    if not k["pareto"]:
        lines.append("  no stops")
    return "\n".join(lines)


# ---------------------------------------------------------------- main
log_dir = find_log_dir()
parts = read_csv(os.path.join(log_dir, "kuka_cell_log.csv"))
events = read_csv(os.path.join(log_dir, "kuka_cell_events.csv"))

if parts and "order" not in parts[0]:
    raise Exception("Old log format. Run the new main_cycle first.")

order = parts[-1]["order"] if (ONLY_LAST_ORDER and parts) else "ALL"
if ONLY_LAST_ORDER:
    parts = [p for p in parts if p["order"] == order]
    events = [e for e in events if e.get("order") == order]

kpi = compute(parts, events)
report = fmt_report(order, kpi)
print(report)

out = os.path.join(log_dir, "kpi_report.txt")
with open(out, "w") as f:
    f.write(report + "\n")

try:
    from robodk.robolink import Robolink
    Robolink().ShowMessage(report + f"\n\nSaved: {out}", True)
except Exception:
    pass

--- Python program dashboard ---
# =====================================================================
#  dashboard.py  -  STEP 3: visual MES dashboard of the KUKA cell
#
#  Reads kuka_cell_log.csv + kuka_cell_events.csv, computes the KPIs
#  (same formulas as kpi_report.py) and writes ONE self-contained file:
#      dashboard.html   (opens in your web browser, no internet needed)
#
#  Run it from RoboDK (Python program, double-click) or: python dashboard.py
# =====================================================================
import csv
import html
import math
import os
import webbrowser
from collections import defaultdict
from datetime import datetime

ONLY_LAST_ORDER = True      # True = last production order only
IDEAL_CYCLE_S = None        # target cycle time (s). None = best cycle observed
LAST_PARTS_ROWS = 15        # rows in the "last parts" table


# ---------------------------------------------------------------- data
def find_log_dir():
    candidates = []
    try:
        from robodk.robolink import Robolink
        d = Robolink().getParam('PATH_OPENSTATION')
        if d:
            candidates.append(str(d))
    except Exception:
        pass
    home = os.path.expanduser("~")
    candidates += [os.path.dirname(os.path.abspath(__file__)),
                   os.path.join(home, "Documents", "KUKA_Cell_MES")]
    for c in candidates:
        if os.path.exists(os.path.join(c, "kuka_cell_log.csv")):
            return c
    for root in [os.path.join(home, d) for d in ("Documents", "OneDrive", "Downloads", "Desktop")]:
        if not os.path.isdir(root):
            continue
        base = root.count(os.sep)
        for folder, subdirs, files in os.walk(root):
            if folder.count(os.sep) - base > 4:
                subdirs[:] = []
                continue
            if "kuka_cell_log.csv" in files:
                return folder
    raise Exception("kuka_cell_log.csv not found. Run main_cycle first.")


def read_csv(path):
    if not os.path.exists(path):
        return []
    with open(path, newline="") as f:
        return list(csv.DictReader(f))


def compute(parts, events):
    n = len(parts)
    n_ok = sum(1 for p in parts if p["result"] == "OK")
    cycles = [float(p["cycle_time_s"]) for p in parts]
    run_time = sum(cycles)
    downtime = sum(float(e["duration_s"]) for e in events)
    planned = run_time + downtime
    ideal = IDEAL_CYCLE_S or min(cycles)
    a = run_time / planned if planned else 0
    p = min(1.0, ideal * n / run_time) if run_time else 0
    q = n_ok / n if n else 0
    pareto = defaultdict(lambda: [0, 0.0])
    for e in events:
        pareto[e["reason"]][0] += 1
        pareto[e["reason"]][1] += float(e["duration_s"])
    pareto = sorted(pareto.items(), key=lambda kv: kv[1][1], reverse=True)
    stops = len(events)
    return dict(n=n, ok=n_ok, nok=n - n_ok, run=run_time, down=downtime, planned=planned,
                ideal=ideal, a=a, p=p, q=q, oee=a * p * q, stops=stops,
                mtbf=run_time / stops if stops else None, mttr=downtime / stops if stops else None,
                avg=run_time / n if n else 0, pareto=pareto)


# ---------------------------------------------------------------- SVG charts
E = html.escape


def cycle_chart(parts, ideal):
    """Vertical bars: cycle time per part + ideal cycle reference line."""
    W, H, L, R, T, B = 1100, 260, 44, 12, 22, 40
    vals = [float(p["cycle_time_s"]) for p in parts]
    vmax = max(10, 10 * math.ceil(max(vals + [ideal]) * 1.1 / 10))   # round axis max to 10
    vmax = vmax if vmax <= 60 else 20 * math.ceil(vmax / 20)
    n = len(vals)
    slot = (W - L - R) / max(n, 1)
    bw = max(4, min(36, slot - 2))
    y = lambda v: T + (H - T - B) * (1 - v / vmax)
    out = [f'<svg viewBox="0 0 {W} {H}" width="{W}" role="img" aria-label="Cycle time per part">']
    step = 10 if vmax <= 60 else (20 if vmax <= 120 else 50)
    for v in range(0, int(vmax) + 1, step):                  # grid + y labels
        out.append(f'<line class="grid" x1="{L}" x2="{W-R}" y1="{y(v):.1f}" y2="{y(v):.1f}"/>')
        out.append(f'<text class="axis" x="{L-6}" y="{y(v)+4:.1f}" text-anchor="end">{v:.0f}</text>')
    for i, (p, v) in enumerate(zip(parts, vals)):
        x = L + i * slot + (slot - bw) / 2
        yy, h = y(v), (H - B) - y(v)
        tip = f'{p["serial"]}: {v:.1f} s ({p["result"]})'
        out.append(f'<g class="hit"><title>{E(tip)}</title>'
                   f'<rect x="{x-1:.1f}" y="{T}" width="{bw+2:.1f}" height="{H-B-T}" fill="transparent"/>'
                   f'<path class="bar" d="M{x:.1f},{H-B} V{yy+4:.1f} Q{x:.1f},{yy:.1f} {x+4:.1f},{yy:.1f} '
                   f'H{x+bw-4:.1f} Q{x+bw:.1f},{yy:.1f} {x+bw:.1f},{yy+4:.1f} V{H-B} Z"/></g>')
        if n <= 15 or i % max(1, n // 10) == 0:
            out.append(f'<text class="axis" x="{x+bw/2:.1f}" y="{H-B+16}" text-anchor="middle">{E(p["serial"][-4:])}</text>')
    yi = y(ideal)
    out.append(f'<line class="ref" x1="{L}" x2="{W-R}" y1="{yi:.1f}" y2="{yi:.1f}"/>')
    out.append(f'<line class="base" x1="{L}" x2="{W-R}" y1="{H-B}" y2="{H-B}"/>')
    out.append(f'<text class="axis" x="{L}" y="{H-4}">serial</text></svg>')
    return "".join(out)


def pareto_chart(pareto, total_down):
    """Horizontal bars: downtime per stop reason, biggest first."""
    if not pareto:
        return '<p class="empty">No stops in this order.</p>'
    W, row, L, R = 520, 34, 170, 100
    H = row * len(pareto) + 8
    vmax = max(sec for _, (c, sec) in pareto) or 1
    out = [f'<svg viewBox="0 0 {W} {H}" width="{W}" role="img" aria-label="Downtime by stop reason">']
    for i, (reason, (count, sec)) in enumerate(pareto):
        yy = 4 + i * row
        w = max(4, (W - L - R) * sec / vmax)
        share = 100 * sec / total_down if total_down else 0
        tip = f"{reason}: {count} stop(s), {sec:.0f} s, {share:.0f} % of downtime"
        out.append(f'<g class="hit"><title>{E(tip)}</title>'
                   f'<rect x="0" y="{yy}" width="{W}" height="{row-4}" fill="transparent"/>'
                   f'<text class="label" x="{L-10}" y="{yy+row/2+2}" text-anchor="end">{E(reason)}</text>'
                   f'<path class="bar" d="M{L},{yy+6} H{L+w-4:.1f} Q{L+w:.1f},{yy+6} {L+w:.1f},{yy+10} '
                   f'V{yy+row-14} Q{L+w:.1f},{yy+row-10} {L+w-4:.1f},{yy+row-10} H{L} Z"/>'
                   f'<text class="value" x="{L+w+8:.1f}" y="{yy+row/2+2}">{sec:.0f} s &middot; {share:.0f} %</text></g>')
    out.append(f'<line class="base" x1="{L}" x2="{L}" y1="0" y2="{H}"/></svg>')
    return "".join(out)


def apq_bars(k):
    rows = [("Availability", k["a"], "running &divide; planned"),
            ("Performance", k["p"], "ideal &times; parts &divide; running"),
            ("Quality", k["q"], "OK &divide; produced")]
    out = []
    for name, v, formula in rows:
        out.append(f'<div class="apq"><div class="apq-head"><span>{name}</span>'
                   f'<strong>{100*v:.1f} %</strong></div>'
                   f'<div class="track"><div class="fill" style="width:{100*v:.1f}%"></div></div>'
                   f'<div class="muted small">{formula}</div></div>')
    return "".join(out)


def status_badge(result):
    if result == "OK":
        return '<span class="badge good">&#10003; OK</span>'
    return '<span class="badge critical">&#10005; NOK</span>'


# ---------------------------------------------------------------- page
def build_html(order, k, parts, events):
    oee = 100 * k["oee"]
    oee_word = "World class" if oee >= 85 else ("Typical plant" if oee >= 60 else "Needs improvement")
    top = k["pareto"][0][0] if k["pareto"] else None
    insight = (f"Biggest loss: <strong>{E(top)}</strong> &mdash; "
               f"{100*k['pareto'][0][1][1]/k['down']:.0f} % of downtime." if top else
               "No stops recorded in this order.")
    rows = []
    for p in reversed(parts[-LAST_PARTS_ROWS:]):
        rows.append(f'<tr><td>{E(p["serial"])}</td><td>{E(p["timestamp"].replace("T", " "))}</td>'
                    f'<td class="num">{float(p["diameter_mm"]):.3f}</td><td>{status_badge(p["result"])}</td>'
                    f'<td class="num">{float(p["cycle_time_s"]):.1f}</td>'
                    f'<td class="num">{float(p.get("downtime_s", 0) or 0):.0f}</td></tr>')
    ev_rows = "".join(f'<tr><td>{E(e["start"].replace("T", " "))}</td><td>{E(e["serial"])}</td>'
                      f'<td>{E(e["station"])}</td><td>{E(e["reason"])}</td>'
                      f'<td class="num">{float(e["duration_s"]):.0f}</td></tr>' for e in reversed(events))
    sec = lambda x: "&ndash;" if x is None else f"{x:.0f} s"
    generated = datetime.now().strftime("%Y-%m-%d %H:%M")

    return f"""<!doctype html>
<html lang="en"><head><meta charset="utf-8">
<meta name="viewport" content="width=device-width, initial-scale=1">
<title>KUKA Cell Dashboard</title>
<style>
:root {{
  color-scheme: light;
  --surface-0:#f4f3f0; --surface-1:#fcfcfb; --border:#e3e2de;
  --text-primary:#0b0b0b; --text-secondary:#52514e; --text-muted:#7a7974;
  --grid:#ecebe7; --series-1:#2a78d6; --track:#ecebe7;
  --good:#0ca30c; --good-text:#006300; --critical:#d03b3b; --critical-text:#b02a2a;
}}
@media (prefers-color-scheme: dark) {{
  :root:where(:not([data-theme="light"])) {{
    color-scheme: dark;
    --surface-0:#121211; --surface-1:#1a1a19; --border:#2e2e2b;
    --text-primary:#ffffff; --text-secondary:#c3c2b7; --text-muted:#8f8e86;
    --grid:#2a2a27; --series-1:#3987e5; --track:#2a2a27;
    --good:#0ca30c; --good-text:#4cc94c; --critical:#d03b3b; --critical-text:#ff8a8a;
  }}
}}
:root[data-theme="dark"] {{
  color-scheme: dark;
  --surface-0:#121211; --surface-1:#1a1a19; --border:#2e2e2b;
  --text-primary:#ffffff; --text-secondary:#c3c2b7; --text-muted:#8f8e86;
  --grid:#2a2a27; --series-1:#3987e5; --track:#2a2a27;
  --good:#0ca30c; --good-text:#4cc94c; --critical:#d03b3b; --critical-text:#ff8a8a;
}}
* {{ box-sizing:border-box; }}
body {{ margin:0; background:var(--surface-0); color:var(--text-primary);
  font:14px/1.45 system-ui,-apple-system,"Segoe UI",Roboto,sans-serif; }}
.wrap {{ max-width:1180px; margin:0 auto; padding:24px 16px 48px; }}
header {{ display:flex; flex-wrap:wrap; justify-content:space-between; align-items:baseline; gap:8px; margin-bottom:18px; }}
h1 {{ font-size:22px; margin:0; }}
h2 {{ font-size:15px; margin:0 0 12px; }}
.muted {{ color:var(--text-secondary); }} .small {{ font-size:12px; }}
.grid2 {{ display:grid; grid-template-columns:repeat(auto-fit,minmax(320px,1fr)); gap:16px; }}
.tiles {{ display:grid; grid-template-columns:repeat(auto-fit,minmax(160px,1fr)); gap:16px; margin-bottom:16px; }}
.card {{ background:var(--surface-1); border:1px solid var(--border); border-radius:12px; padding:18px; min-width:0; }}
.tile .label {{ color:var(--text-secondary); font-size:12px; text-transform:uppercase; letter-spacing:.04em; }}
.tile .big {{ font-size:30px; font-weight:650; margin-top:4px; font-variant-numeric:tabular-nums; }}
.hero .big {{ font-size:clamp(30px,6vw,44px); white-space:nowrap; }}
.tile .big {{ white-space:nowrap; }}
.apq {{ margin-bottom:14px; }}
.apq-head {{ display:flex; justify-content:space-between; margin-bottom:6px; }}
.track {{ height:8px; background:var(--track); border-radius:4px; overflow:hidden; }}
.fill {{ height:100%; background:var(--series-1); border-radius:4px; }}
svg {{ max-width:100%; height:auto; display:block; overflow:visible; }}
svg .grid {{ stroke:var(--grid); stroke-width:1; }}
svg .base {{ stroke:var(--text-muted); stroke-width:1; }}
svg .bar {{ fill:var(--series-1); }}
svg .hit:hover .bar {{ opacity:.8; }}
svg .ref {{ stroke:var(--text-secondary); stroke-width:1.5; }}
svg text {{ font:12px system-ui,-apple-system,"Segoe UI",sans-serif; fill:var(--text-secondary); }}
svg .label {{ fill:var(--text-primary); }}
svg .value, svg .reflabel {{ fill:var(--text-secondary); }}
.insight {{ margin-top:10px; padding:10px 12px; border-left:3px solid var(--series-1); background:var(--surface-0); border-radius:6px; }}
.table-wrap {{ overflow-x:auto; }}
table {{ width:100%; border-collapse:collapse; font-size:13px; }}
th, td {{ text-align:left; padding:8px 10px; border-bottom:1px solid var(--border); white-space:nowrap; }}
th {{ color:var(--text-secondary); font-weight:600; font-size:12px; }}
td.num, th.num {{ text-align:right; font-variant-numeric:tabular-nums; }}
.badge {{ display:inline-block; padding:2px 8px; border-radius:999px; font-size:12px; font-weight:600; }}
.badge.good {{ color:var(--good-text); background:color-mix(in srgb, var(--good) 14%, transparent); }}
.badge.critical {{ color:var(--critical-text); background:color-mix(in srgb, var(--critical) 14%, transparent); }}
.empty {{ color:var(--text-secondary); }}
section {{ margin-top:16px; }}
</style></head>
<body><div class="wrap">
<header>
  <div><h1>KUKA KR 10 machine-tending cell</h1>
  <div class="muted">Production order <strong>{E(order)}</strong> &middot; {k['n']} parts</div></div>
  <div class="muted small">Generated {generated}</div>
</header>

<div class="tiles">
  <div class="card tile hero"><div class="label">OEE</div><div class="big">{oee:.1f} %</div>
    <div class="muted small">{oee_word} (benchmark: world class &ge; 85 %)</div></div>
  <div class="card tile"><div class="label">Good parts</div><div class="big">{k['ok']} / {k['n']}</div>
    <div class="small">{status_badge('OK')} {k['ok']} &nbsp; {status_badge('NOK')} {k['nok']}</div></div>
  <div class="card tile"><div class="label">Avg cycle time</div><div class="big">{k['avg']:.1f} s</div>
    <div class="muted small">ideal {k['ideal']:.1f} s</div></div>
  <div class="card tile"><div class="label">Downtime</div><div class="big">{k['down']:.0f} s</div>
    <div class="muted small">{k['stops']} stop{'s' if k['stops'] != 1 else ''} &middot; MTBF {sec(k['mtbf'])} &middot; MTTR {sec(k['mttr'])}</div></div>
</div>

<div class="grid2">
  <div class="card"><h2>OEE = Availability &times; Performance &times; Quality</h2>{apq_bars(k)}
    <div class="insight">{insight}</div></div>
  <div class="card"><h2>Downtime by stop reason (Pareto)</h2>{pareto_chart(k['pareto'], k['down'])}</div>
</div>

<section class="card"><h2>Cycle time per part (s)</h2>{cycle_chart(parts, k['ideal'])}
  <div class="muted small">Hover a bar for details. Horizontal line = ideal cycle time ({k['ideal']:.1f} s).</div></section>

<div class="grid2">
<section class="card"><h2>Last parts (traceability)</h2><div class="table-wrap"><table>
<thead><tr><th>Serial</th><th>Time</th><th class="num">&Oslash; (mm)</th><th>Result</th><th class="num">Cycle (s)</th><th class="num">Stop (s)</th></tr></thead>
<tbody>{''.join(rows)}</tbody></table></div></section>
<section class="card"><h2>Stop events</h2><div class="table-wrap"><table>
<thead><tr><th>Start</th><th>Serial</th><th>Station</th><th>Reason</th><th class="num">Duration (s)</th></tr></thead>
<tbody>{ev_rows or '<tr><td colspan="5" class="empty">No stops</td></tr>'}</tbody></table></div></section>
</div>
</div></body></html>"""


# ---------------------------------------------------------------- main
log_dir = find_log_dir()
parts = read_csv(os.path.join(log_dir, "kuka_cell_log.csv"))
events = read_csv(os.path.join(log_dir, "kuka_cell_events.csv"))
if not parts:
    raise Exception("No parts in kuka_cell_log.csv. Run main_cycle first.")
if "order" not in parts[0]:
    raise Exception("Old log format. Run the new main_cycle first.")

order = parts[-1]["order"] if ONLY_LAST_ORDER else "ALL"
if ONLY_LAST_ORDER:
    parts = [p for p in parts if p["order"] == order]
    events = [e for e in events if e.get("order") == order]

kpi = compute(parts, events)
out = os.path.join(log_dir, "dashboard.html")
with open(out, "w", encoding="utf-8") as f:
    f.write(build_html(order, kpi, parts, events))
print(f"Dashboard written: {out}")
webbrowser.open("file:///" + out.replace("\\", "/"))
